(* IEC 61131-3 sources: machine-design-framework/examples/pick-glue-place-broken/plc/generated, 2 files *)

(* ---- GVL_Cycle.st ---- *)
(* GENERATED from cycle.yaml - DO NOT EDIT. source-hash: d747394b20adf07e *)
(* Commanded angles (deg). Effective timing = commanded + device delay; see GLUE-BEAD/PROD-* checks. *)
VAR_GLOBAL CONSTANT
    VACUUM_ON  : REAL := 10.0000;
    VACUUM_OFF : REAL := 222.0000;
    GLUE_GUN_ON  : REAL := 128.6400;
    GLUE_GUN_OFF : REAL := 130.4000;
    VAC_OK_CHECK : REAL := 26.0000;
    DOUBLE_SHEET_CHECK : REAL := 75.0000;
    PARK_ANGLE : REAL := 355.0000;
END_VAR

(* ---- GVL_IO.st ---- *)
(* GENERATED from io_list.yaml - DO NOT EDIT. source-hash: 5f45f90c360e175b *)
VAR_GLOBAL
    rAngle : REAL;   (* in  virtual *)
    xMasterRun : BOOL;   (* out  virtual *)
    xVacuum : BOOL;   (* out  DO1.0 VAC_VALVE *)
    xGlueGun : BOOL;   (* out  DO1.1 GLUE_VALVE *)
    xLampFault : BOOL;   (* out  DO1.2 LAMP_FAULT *)
    xVacOk : BOOL;   (* in  DI1.0 VAC_SWITCH *)
    xDoubleSheet : BOOL;   (* in  DI1.1 DOUBLE_SENSOR *)
    xAirOk : BOOL;   (* in  DI1.2 AIR_SWITCH *)
    xGlueReady : BOOL;   (* in  DI1.3 GLUE_UNIT *)
    xStartPb : BOOL;   (* in  DI1.4 OP_PANEL *)
    xStopPb : BOOL;   (* in  DI1.5 OP_PANEL *)
    xResetPb : BOOL;   (* in  DI1.6 OP_PANEL *)
    xGuardClosed : BOOL;   (* in  SDI1.0 GUARD_SWITCH *)
    xEStopOk : BOOL;   (* in  SDI1.1 ESTOP *)
END_VAR
